Staubli VAL3: main.pgx

public program main()
begin
  if rs:sPageUsing!="main"
    rs:sPageUsing="main"
    //
    call util:loadingPage()
    //
    userPage(rs:sPageUsing)
    delay(1)
  endIf
end
